(* IEC 61131-3 sources: plcassist-cli/packages/volt-lsp-iec/test-corpus/awa-palletizer/Device/Plc Logic/Application/Library Manager/(unresolved)/cmpopcuaserver interfaces, 1 file *)

(* ---- EVENTIDS.gvl ---- *)
VAR_GLOBAL
	CMPID_CMPOPCUASERVER : DWORD := 16#124;
	EVTPARAMID_CMPOPCUASERVERSESSIONSCHANGED : WORD := 16#1;
	EVTVERSION_CMPOPCUASERVERSESSIONSCHANGED : WORD := 16#1;
	EVT_CMPOPCUASERVERSESSIONSCHANGED : DWORD := (SHL(UINT_TO_DWORD(EventClass.EVTCLASS_INFO), 16) OR 16#1);
END_VAR
